FUNCTION_BLOCK basicDesinfeccao (* Logica da desinfeccao (limitacao de vazao pela 700-VC-01, totalizacao, alarmes) *)
  (* Standard: 61499-2 *)
  (* Version 1.1, 12/11/2026, Hidryco, Hidryco, 1.1: sentido dos disjuntores conferido em campo - PCE/PCM: 1 = ligado (invertido); UV-01/02, VC-01 e monovia: 1 = ligado (sem mudanca); variaveis e tags sem mudanca de nome; alarme de disjuntor desativado (stsAvisoDisjuntor sempre FALSE), status dos disjuntores mantidos. 1.0: PID continuo sobre a 700-FT-01 (m3/h) comandando a 700-VC-01; FT em falha ou valvula indisponivel mantem a posicao; totalizador persistente; vazao alta e variacao brusca *)
  PACKAGE Hidryco.HidrycoLib;
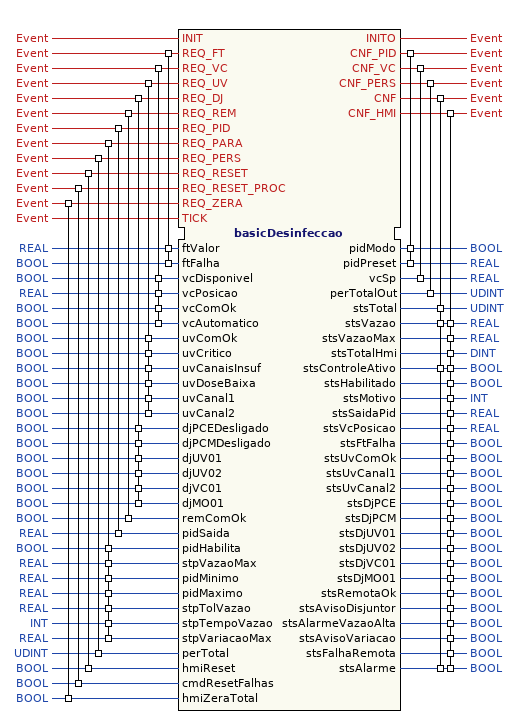
  EVENT_INPUT
    INIT; (* Inicializacao *)
    REQ_FT WITH ftValor, ftFalha; (* 700-FT-01 (Parshall) *)
    REQ_VC WITH vcDisponivel, vcPosicao, vcComOk, vcAutomatico; (* 700-VC-01 *)
    REQ_UV WITH uvComOk, uvCritico, uvCanaisInsuf, uvDoseBaixa, uvCanal1, uvCanal2; (* 700-UV-01/02 *)
    REQ_DJ WITH djPCEDesligado, djPCMDesligado, djUV01, djUV02, djVC01, djMO01; (* Disjuntores (remota da desinfeccao) *)
    REQ_REM WITH remComOk; (* Remota da desinfeccao comunicando (COM_OK do IO_DI32) *)
    REQ_PID WITH pidSaida; (* Saida do PID *)
    REQ_PARA WITH pidHabilita, stpVazaoMax, pidMinimo, pidMaximo, stpTolVazao, stpTempoVazao, stpVariacaoMax; (* IHM: parametros *)
    REQ_PERS WITH perTotal; (* Totalizador lido da persistencia *)
    REQ_RESET WITH hmiReset; (* IHM: reset *)
    REQ_RESET_PROC WITH cmdResetFalhas; (* Processo: reset *)
    REQ_ZERA WITH hmiZeraTotal; (* IHM: zera o totalizador *)
    TICK; (* Base de tempo de 1 s *)
  END_EVENT
  EVENT_OUTPUT
    INITO; (* Inicializacao concluida *)
    CNF_PID WITH pidModo, pidPreset; (* Modo do pidCtl (automatico ou tracking da posicao) *)
    CNF_VC WITH vcSp; (* Posicao pedida a 700-VC-01 *)
    CNF_PERS WITH perTotalOut; (* Grava o totalizador *)
    CNF WITH stsVazao, stsTotal, stsControleAtivo, stsAlarme; (* Status para o processo *)
    CNF_HMI WITH stsVazao, stsVazaoMax, stsTotalHmi, stsControleAtivo, stsHabilitado, stsMotivo, stsSaidaPid, stsVcPosicao, stsFtFalha, stsUvComOk, stsUvCanal1, stsUvCanal2, stsDjPCE, stsDjPCM, stsDjUV01, stsDjUV02, stsDjVC01, stsDjMO01, stsRemotaOk, stsAvisoDisjuntor, stsAlarmeVazaoAlta, stsAvisoVariacao, stsFalhaRemota, stsAlarme; (* Status para a IHM e alarmes *)
  END_EVENT
  VAR_INPUT
    ftValor : REAL; (* Vazao 700-FT-01 (m3/h) *)
    ftFalha : BOOL; (* 700-FT-01 com sinal em falha *)
    vcDisponivel : BOOL; (* VC-01 disponivel para o automatico *)
    vcPosicao : REAL; (* Posicao da VC-01 (%) *)
    vcComOk : BOOL; (* VC-01 comunicando *)
    vcAutomatico : BOOL; (* VC-01 em automatico *)
    uvComOk : BOOL;
    uvCritico : BOOL;
    uvCanaisInsuf : BOOL;
    uvDoseBaixa : BOOL;
    uvCanal1 : BOOL;
    uvCanal2 : BOOL;
    djPCEDesligado : BOOL; (* Remota %I0.0 *)
    djPCMDesligado : BOOL; (* Remota %I0.1 *)
    djUV01 : BOOL; (* Remota %I0.2 *)
    djUV02 : BOOL; (* Remota %I0.3 *)
    djVC01 : BOOL; (* Remota %I0.4 *)
    djMO01 : BOOL; (* Remota %I0.5 *)
    remComOk : BOOL; (* Remota comunicando (COM_OK publicado pelo IO_DI32 da remota) *)
    pidSaida : REAL; (* Saida do PID (%) *)
    pidHabilita : BOOL; (* Controle de vazao habilitado *)
    stpVazaoMax : REAL; (* Vazao maxima de lancamento (m3/h) *)
    pidMinimo : REAL; (* Saida minima do PID (%) *)
    pidMaximo : REAL; (* Saida maxima do PID (%) *)
    stpTolVazao : REAL; (* Tolerancia acima do limite para o alarme (%) *)
    stpTempoVazao : INT; (* Tempo acima do limite para o alarme (s); 0 = desligado *)
    stpVariacaoMax : REAL; (* Variacao maxima da vazao em 1 min (m3/h); 0 = desligado *)
    perTotal : UDINT; (* Totalizador persistido (m3) *)
    hmiReset : BOOL;
    cmdResetFalhas : BOOL;
    hmiZeraTotal : BOOL;
  END_VAR
  VAR_OUTPUT
    pidModo : BOOL; (* TRUE = PID em automatico; FALSE = saida segue a posicao da valvula *)
    pidPreset : REAL; (* Valor de tracking do PID (posicao da valvula) *)
    vcSp : REAL; (* Posicao pedida a 700-VC-01 (%) *)
    perTotalOut : UDINT; (* Totalizador a gravar (m3) *)
    stsTotal : UDINT; (* Volume totalizado (m3) *)
    stsVazao : REAL; (* Vazao do efluente final 700-FT-01 (m3/h) *)
    stsVazaoMax : REAL; (* Vazao maxima de lancamento em uso (m3/h) *)
    stsTotalHmi : DINT; (* Volume totalizado (m3) *)
    stsControleAtivo : BOOL; (* PID controlando a 700-VC-01 *)
    stsHabilitado : BOOL; (* Controle de vazao habilitado pelo operador *)
    stsMotivo : INT; (* Controle: 0 controlando, 1 desabilitado, 2 FT-01 em falha, 3 valvula indisponivel, 4 retomando (3 s) *)
    stsSaidaPid : REAL; (* Saida do PID (%) *)
    stsVcPosicao : REAL; (* Posicao da 700-VC-01 (%) *)
    stsFtFalha : BOOL; (* 700-FT-01 em falha *)
    stsUvComOk : BOOL; (* UV comunicando *)
    stsUvCanal1 : BOOL; (* UV canal 1 operando *)
    stsUvCanal2 : BOOL; (* UV canal 2 operando *)
    stsDjPCE : BOOL; (* Remota %I0.0: disjuntor desligado PCE *)
    stsDjPCM : BOOL; (* Remota %I0.1: disjuntor desligado PCM desinfeccao *)
    stsDjUV01 : BOOL; (* Remota %I0.2: disjuntor ligado 700-UV-01 *)
    stsDjUV02 : BOOL; (* Remota %I0.3: disjuntor ligado 700-UV-02 *)
    stsDjVC01 : BOOL; (* Remota %I0.4: disjuntor ligado 700-VC-01 *)
    stsDjMO01 : BOOL; (* Remota %I0.5: disjuntor ligado 700-MO-01 (monovia) *)
    stsRemotaOk : BOOL; (* Remota da desinfeccao comunicando *)
    stsAvisoDisjuntor : BOOL; (* Disjuntor do PCE, PCM, UV ou VC-01 desligado *)
    stsAlarmeVazaoAlta : BOOL; (* Vazao acima do limite de lancamento (memorizado) *)
    stsAvisoVariacao : BOOL; (* Variacao brusca da vazao de lancamento (memorizado) *)
    stsFalhaRemota : BOOL; (* Falha de comunicacao com a remota da desinfeccao *)
    stsAlarme : BOOL; (* Algum alarme da desinfeccao *)
  END_VAR
  VAR
    initDone : BOOL;
    primeiro : BOOL := TRUE;
    acc : REAL; (* Fracao do totalizador (m3) *)
    nInteiro : UDINT;
    tGrava : INT;
    totalGravado : UDINT;
    persLido : BOOL;
    tAlta : INT;
    tVar : INT;
    qAnt : REAL;
    qAntOk : BOOL;
    oldModo : BOOL;
    oldSp : REAL := -100.0;
    oldSig : INT := -1;
    sig : INT;
    rLimite : REAL;
    condOk : BOOL;
    tEstavel : INT; (* Segundos com as condicoes do controle OK *)
  END_VAR
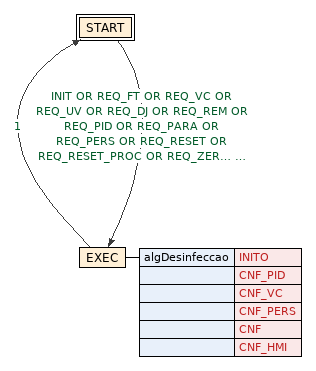
  EC_STATES
    START; (* Estado inicial *)
    EXEC : algDesinfeccao -> INITO, -> CNF_PID, -> CNF_VC, -> CNF_PERS, -> CNF, -> CNF_HMI; (* Executa a logica; o algoritmo decide quais eventos saem *)
  END_STATES
  EC_TRANSITIONS
    START TO EXEC := INIT OR REQ_FT OR REQ_VC OR REQ_UV OR REQ_DJ OR REQ_REM OR REQ_PID OR REQ_PARA OR REQ_PERS OR REQ_RESET OR REQ_RESET_PROC OR REQ_ZERA OR TICK;
    EXEC TO START := 1;
  END_TRANSITIONS
  ALGORITHM algDesinfeccao IN ST: (* Logica completa (um unico algoritmo) *)
(* =====================================================================
   basicDesinfeccao v1.0 - logica do CAT Desinfeccao_UV (HidrycoLib)
   Limitacao da vazao de lancamento pela 700-VC-01 (borboleta DN600 na
   saida do tanque de amortecimento) com PID continuo sobre a 700-FT-01
   (Parshall, m3/h) - manual REL-007 2.4.1: maximo 345 L/s = 1242 m3/h.
   Regras (definidas pelo usuario):
   - PID continuo; valvula modulante (Valvula_Coester cfgModulante);
   - FT-01 em falha, PID desabilitado ou valvula indisponivel: a valvula
     mantem a posicao (referencia = posicao medida) e o PID acompanha a
     posicao (tracking) para retomar sem salto;
   - totalizacao em m3 (persistente); alarme de vazao acima do limite e
     aviso de variacao brusca (manual 2.4.4), ambos ate o reset;
   - o UV (Trojan) e somente monitorado: nao ha comando do CLP.
   ===================================================================== *)

INITO    := FALSE;
CNF_PID  := FALSE;
CNF_VC   := FALSE;
CNF_PERS := FALSE;
CNF      := FALSE;
CNF_HMI  := FALSE;

IF INIT THEN
    initDone := TRUE;
    INITO := TRUE;
END_IF;
IF NOT initDone THEN
    RETURN;
END_IF;

(* ---- 1. Totalizador persistente ---- *)
IF REQ_PERS AND NOT persLido THEN
    persLido := TRUE;
    IF perTotal > stsTotal THEN
        stsTotal := perTotal;
    END_IF;
    totalGravado := stsTotal;
END_IF;
IF REQ_ZERA AND hmiZeraTotal THEN
    stsTotal := 0;
    acc := 0.0;
    CNF_PERS := TRUE;
END_IF;
IF TICK AND NOT ftFalha AND (ftValor > 0.0) THEN
    acc := acc + ftValor / 3600.0;
    IF acc >= 1.0 THEN
        nInteiro := REAL_TO_UDINT(acc - 0.5);
        stsTotal := stsTotal + nInteiro;
        acc := acc - UDINT_TO_REAL(nInteiro);
    END_IF;
END_IF;
IF TICK THEN
    tGrava := tGrava + 1;
    IF (tGrava >= 60) AND (stsTotal <> totalGravado) THEN
        tGrava := 0;
        CNF_PERS := TRUE;
    END_IF;
END_IF;
IF CNF_PERS THEN
    perTotalOut := stsTotal;
    totalGravado := stsTotal;
END_IF;
stsTotalHmi := UDINT_TO_DINT(stsTotal);

(* ---- 2. Controle da 700-VC-01 ---- *)
stsVazao := ftValor;
stsFtFalha := ftFalha;
stsHabilitado := pidHabilita;
stsVazaoMax := stpVazaoMax;
stsVcPosicao := vcPosicao;
stsSaidaPid := pidSaida;
(* o controle so (re)assume com tudo OK ha 3 s: o PID acompanha a posicao com o PV ja valido e volta sem salto *)
condOk := pidHabilita AND NOT ftFalha AND vcDisponivel;
IF NOT condOk THEN
    tEstavel := 0;
ELSIF TICK AND (tEstavel < 3) THEN
    tEstavel := tEstavel + 1;
END_IF;
IF NOT pidHabilita THEN
    stsMotivo := 1;
ELSIF ftFalha THEN
    stsMotivo := 2;
ELSIF NOT vcDisponivel THEN
    stsMotivo := 3;
ELSIF tEstavel < 3 THEN
    stsMotivo := 4;
ELSE
    stsMotivo := 0;
END_IF;
stsControleAtivo := stsMotivo = 0;
pidModo := stsControleAtivo;
pidPreset := vcPosicao;
IF stsControleAtivo THEN
    vcSp := LIMIT(pidMinimo, pidSaida, pidMaximo);
ELSE
    vcSp := vcPosicao;                     (* mantem a posicao *)
END_IF;
IF primeiro OR (pidModo <> oldModo) OR REQ_VC THEN
    CNF_PID := TRUE;
    oldModo := pidModo;
END_IF;
IF primeiro OR TICK OR (ABS(vcSp - oldSp) >= 0.5) THEN
    CNF_VC := TRUE;
    oldSp := vcSp;
END_IF;

(* ---- 3. Alarmes de processo ---- *)
IF (REQ_RESET AND hmiReset) OR (REQ_RESET_PROC AND cmdResetFalhas) THEN
    stsAlarmeVazaoAlta := FALSE;
    stsAvisoVariacao := FALSE;
    tAlta := 0;
END_IF;
rLimite := stpVazaoMax * (1.0 + stpTolVazao / 100.0);
IF TICK THEN
    IF (stpTempoVazao > 0) AND NOT ftFalha AND (stpVazaoMax > 0.0) AND (ftValor > rLimite) THEN
        tAlta := tAlta + 1;
        IF tAlta >= stpTempoVazao THEN
            stsAlarmeVazaoAlta := TRUE;
        END_IF;
    ELSE
        tAlta := 0;
    END_IF;
    tVar := tVar + 1;
    IF tVar >= 60 THEN
        tVar := 0;
        IF qAntOk AND NOT ftFalha AND (stpVariacaoMax > 0.0) AND (ABS(ftValor - qAnt) > stpVariacaoMax) THEN
            stsAvisoVariacao := TRUE;
        END_IF;
        qAnt := ftValor;
        qAntOk := NOT ftFalha;
    END_IF;
END_IF;
stsRemotaOk := remComOk;
stsFalhaRemota := NOT stsRemotaOk;
IF stsRemotaOk THEN
    (* sentido conferido em campo (12/11/2026): %I0.0 PCE e %I0.1 PCM = 1 com o disjuntor LIGADO
       (invertido em relacao ao nome); %I0.2 a %I0.5 (UV-01, UV-02, VC-01, monovia) = 1 ligado.
       Nomes das variaveis/tags mantidos. *)
    stsDjPCE := NOT djPCEDesligado; stsDjPCM := NOT djPCMDesligado;
    stsDjUV01 := djUV01; stsDjUV02 := djUV02; stsDjVC01 := djVC01; stsDjMO01 := djMO01;
    stsAvisoDisjuntor := FALSE;   (* alarme de disjuntor desativado a pedido do usuario (12/11/2026); os status continuam *)
ELSE
    stsAvisoDisjuntor := FALSE;
END_IF;
stsUvComOk := uvComOk;
stsUvCanal1 := uvCanal1;
stsUvCanal2 := uvCanal2;
stsAlarme := stsAlarmeVazaoAlta OR stsAvisoVariacao OR stsAvisoDisjuntor OR stsFalhaRemota OR ftFalha;

(* ---- 4. Eventos ---- *)
sig := stsMotivo;
IF stsAlarmeVazaoAlta THEN sig := sig + 8; END_IF;
IF stsAvisoVariacao THEN sig := sig + 16; END_IF;
IF stsAvisoDisjuntor THEN sig := sig + 32; END_IF;
IF stsFalhaRemota THEN sig := sig + 64; END_IF;
IF stsAlarme THEN sig := sig + 128; END_IF;
IF primeiro OR TICK OR REQ_PARA OR REQ_RESET OR REQ_ZERA OR (sig <> oldSig) THEN
    CNF_HMI := TRUE;
END_IF;
IF primeiro OR TICK OR (sig <> oldSig) THEN
    CNF := TRUE;
END_IF;
oldSig := sig;
primeiro := FALSE;
  END_ALGORITHM
END_FUNCTION_BLOCK
